Staubli VAL3: progTemplate.pjx

--- progTemplate.pjx ---
Parameters version=s8.12.1Cs9_BS2449 stackSize=5000 millimeterUnit=true
Program file=start.pgx
Program file=stop.pgx
Data file=progTemplate.dtx
Type name=ifItem path=Disk://source/template/ifItem/ifItem.pjx
Type name=switchItem path=Disk://source/template/switchItem/switchItem.pjx
Type name=forItem path=Disk://source/template/forItem/forItem.pjx

--- progTemplate.dtx ---
public string sTRAJname
public num nType
public ifItem iIfItem
  [0]
    num nSigType[3]
    num nSigIndex[3]
    num nValue[3]
    bool bANDOR[2]
public switchItem sSwitchItem
  [0]
    num nSwitchValue
    string sIOValue
    bool bIOdisable
public forItem fForItem
  [0]
    num nLoopValue
    bool bIOdisable
    string sIOindex
    string sForTRAJ

--- start.pgx ---
program start()
begin
end

--- stop.pgx ---
program stop()
begin
end
